{attribute 'TcGvlVarFlags' := 'OPC'}
VAR_GLOBAL
    // Commands — written by Python over ADS, sent to device every cycle
    // ADS symbol: GVL_UartBridge.stCmd
    stCmd               : ST_UartBridgeCmd;

    // Status — read from device every cycle, read by Python over ADS
    // ADS symbol: GVL_UartBridge.stStatus
    stStatus            : ST_UartBridgeStatus;
END_VAR

(* stored: Version 1.1.0.1, ProductVersion 3.1.4026.18
   GVL GVL_UartBridge: Id {c80e02e1-177b-4ccb-89b2-7fafc7a9d400} *)
